(* IEC 61131-3 sources: OpenUnit/plc/projects/GEN/pous/function-blocks, 7 files *)

(* ---- FB_LOOP.st ---- *)
(* PID loop bound to its faceplate tags (<loop>_PV/_SP/_OUT/_MODE/_KP/_TI/_TD/_CSP/_STS).
   Ideal (ISA) PID working in % of span, back-calculation anti-windup, derivative on
   measurement with a 0.1*TD filter, feed-forward and bumpless MAN/AUTO/CAS transfer.
   MODE: 0 MAN, 1 AUTO, 2 CAS.  STS bits: 1 interlock, 2 tracking, 4 high limit, 8 low limit,
   16 cascade setpoint available.  Mirrors Loop + PID in the JavaScript controller runtime. *)
FUNCTION_BLOCK FB_LOOP
  VAR_INPUT
    PV_IN : REAL;              (* process value, engineering units *)
    CSP_IN : REAL;             (* cascade / remote setpoint *)
    CSP_OK : BOOL;             (* remote setpoint supplied and available *)
    FF : REAL;                 (* feed-forward, output engineering units *)
    FORCE_MAN : BOOL;          (* interlock: force manual *)
    TRK : BOOL;                (* track TRK_VAL *)
    TRK_VAL : REAL;
    OUT_HI : REAL := 1.0E30;   (* dynamic output limits, engineering units *)
    OUT_LO : REAL := -1.0E30;
    SP_LO : REAL := -1.0E30;
    SP_HI : REAL := 1.0E30;
    DTS : REAL;                (* simulation time step, s *)
    RESYNC : BOOL;             (* first scan after start-up / initial condition *)
    PV_MIN : REAL := 0.0;      (* configuration from the register map *)
    PV_MAX : REAL := 100.0;
    OUT_MIN : REAL := 0.0;
    OUT_MAX : REAL := 100.0;
    DIRECT : BOOL;             (* direct acting: output rises when PV > SP *)
    SP_TRACK : BOOL := TRUE;   (* setpoint tracks PV in manual *)
    CAS_CFG : BOOL;            (* loop has a cascade input *)
    REF_DT : REAL;             (* > 0: detune when the step exceeds REF_DT (fast time) *)
  END_VAR
  VAR_IN_OUT
    SP : REAL;
    OUT : REAL;
    MODE : DINT;
    KP : REAL;
    TI : REAL;
    TD : REAL;
    PV : REAL;
    CSP : REAL;
    STS : DINT;
  END_VAR
  VAR_OUTPUT
    Q : REAL;                  (* output, engineering units *)
    AUTO : BOOL;               (* not in manual *)
  END_VAR
  VAR
    integ : REAL;
    outPct : REAL;
    prevPv : REAL;
    havePrev : BOOL;
    dState : REAL;
    lastMode : DINT;
    wasTracking : BOOL;
    slow : REAL;
    kpE : REAL;
    tiE : REAL;
    tdE : REAL;
    m : DINT;
    stsW : DINT;
    casOk : BOOL;
    spv : REAL;
    spanO : REAL;
    spanP : REAL;
    ffPct : REAL;
    hiPct : REAL;
    loPct : REAL;
    err : REAL;
    trkPct : REAL;
    p : REAL;
    d : REAL;
    dpv : REAL;
    raw : REAL;
    alpha : REAL;
    hi : REAL;
    lo : REAL;
    unc : REAL;
    doTrack : BOOL;
  END_VAR

  slow := 1.0;
  IF REF_DT > 0.0 AND DTS > REF_DT THEN
    slow := REF_DT / DTS;
  END_IF;
  kpE := MAX(0.0, KP) * slow;
  tiE := MAX(0.0, TI) / slow;
  tdE := MAX(0.0, TD);

  m := MODE;
  IF m > 2 OR m < 0 THEN
    m := 0;
  END_IF;
  stsW := 0;
  IF FORCE_MAN THEN
    m := 0;
    stsW := stsW + 1;
  END_IF;
  casOk := CAS_CFG AND CSP_OK;
  IF casOk THEN
    stsW := stsW + 16;
  END_IF;
  IF m = 2 AND NOT casOk THEN
    m := 1;
  END_IF;
  spv := SP;
  IF m = 2 THEN
    spv := CSP_IN;
  END_IF;
  spv := LIMIT(SP_LO, spv, SP_HI);

  spanO := OUT_MAX - OUT_MIN;
  IF spanO = 0.0 THEN
    spanO := 1.0;
  END_IF;
  spanP := PV_MAX - PV_MIN;
  IF spanP = 0.0 THEN
    spanP := 1.0;
  END_IF;
  ffPct := FF / spanO * 100.0;
  hiPct := 100.0;
  IF OUT_HI < 1.0E29 THEN
    hiPct := (MIN(OUT_HI, OUT_MAX) - OUT_MIN) / spanO * 100.0;
  END_IF;
  loPct := 0.0;
  IF OUT_LO > -1.0E29 THEN
    loPct := (MAX(OUT_LO, OUT_MIN) - OUT_MIN) / spanO * 100.0;
  END_IF;
  err := (spv - PV_IN) / spanP * 100.0;
  IF DIRECT THEN
    err := -err;
  END_IF;

  (* Tracking / manual: force the output and back-calculate the integrator *)
  doTrack := FALSE;
  IF TRK THEN
    trkPct := (TRK_VAL - OUT_MIN) / spanO * 100.0;
    doTrack := TRUE;
    stsW := stsW + 2;
  ELSIF m = 0 THEN
    trkPct := LIMIT(loPct, (OUT - OUT_MIN) / spanO * 100.0, hiPct);
    doTrack := TRUE;
  ELSIF RESYNC OR lastMode = 0 OR wasTracking THEN
    trkPct := (OUT - OUT_MIN) / spanO * 100.0;
    doTrack := TRUE;
  END_IF;
  IF doTrack THEN
    outPct := LIMIT(0.0, trkPct, 100.0);
    integ := outPct - kpE * err - ffPct;
    prevPv := PV_IN;
    havePrev := TRUE;
    dState := 0.0;
  END_IF;

  IF TRK THEN
    IF m = 0 AND SP_TRACK THEN
      spv := PV_IN;
    END_IF;
  ELSIF m = 0 THEN
    IF SP_TRACK THEN
      spv := LIMIT(SP_LO, PV_IN, SP_HI);
    END_IF;
  ELSE
    (* Automatic: PID update *)
    IF DTS > 0.0 THEN
      p := kpE * err;
      IF tiE > 0.0 THEN
        integ := integ + kpE * err * DTS / tiE;
      END_IF;
      d := 0.0;
      IF tdE > 0.0 AND havePrev THEN
        dpv := ((PV_IN - prevPv) / spanP * 100.0) / DTS;
        IF DIRECT THEN
          raw := kpE * tdE * dpv;
        ELSE
          raw := -kpE * tdE * dpv;
        END_IF;
        alpha := DTS / (0.1 * tdE + DTS);
        dState := dState + alpha * (raw - dState);
        d := dState;
      END_IF;
      prevPv := PV_IN;
      havePrev := TRUE;
      hi := MIN(hiPct, 100.0);
      lo := MAX(loPct, 0.0);
      unc := p + integ + d + ffPct;
      outPct := LIMIT(lo, unc, hi);
      IF unc <> outPct THEN
        integ := outPct - p - d - ffPct;
      END_IF;
      IF tiE <= 0.0 THEN
        integ := LIMIT(-1.0E6, integ, 1.0E6);
      END_IF;
    END_IF;
    IF outPct >= hiPct - 0.000001 THEN
      stsW := stsW + 4;
    END_IF;
    IF outPct <= loPct + 0.000001 THEN
      stsW := stsW + 8;
    END_IF;
  END_IF;

  wasTracking := TRK;
  Q := OUT_MIN + outPct / 100.0 * spanO;
  PV := PV_IN;
  SP := spv;
  OUT := Q;
  MODE := m;
  IF CSP_OK THEN
    CSP := CSP_IN;
  ELSE
    CSP := spv;
  END_IF;
  STS := stsW;
  lastMode := m;
  AUTO := m <> 0;
END_FUNCTION_BLOCK

(* ---- FB_MOTOR.st ---- *)
(* Motor / pump / fan device block.  Drives the field command from START/STOP pulses
   (cleared after use), auto start/stop logic and the protective interlock.  A trip of the
   drive is latched (TRIP) until the operator presses STOP, so a standby unit can start on it.
   SYNC (initial condition) aligns the command with the running feedback.  CMD_SET forces the
   command from a sequence, like an operator start without the permissive check. *)
FUNCTION_BLOCK FB_MOTOR
  VAR_INPUT
    RUN_FB : BOOL;             (* field: running *)
    TRIP_FB : BOOL;            (* field: tripped *)
    PERMIT : BOOL := TRUE;     (* start permissive *)
    ILK : BOOL;                (* protective interlock (stops and blocks) *)
    AUTO_START : BOOL;
    AUTO_STOP : BOOL;
    SYNC : BOOL;
    CMD_SET : BOOL;
    CMD_VAL : BOOL;
  END_VAR
  VAR_IN_OUT
    START : BOOL;              (* operator pulse *)
    STOP : BOOL;               (* operator pulse *)
    MODE : DINT;               (* 0 MAN, 1 AUTO / standby *)
    CMD : BOOL;                (* field command *)
    RUN : BOOL;
    TRIP : BOOL;
    PERM : BOOL;
    ILK_T : BOOL;
  END_VAR
  VAR_OUTPUT
    RUNNING : BOOL;
    LATCHED : BOOL;            (* trip latch (cleared by STOP) *)
    TRIPPED : BOOL;            (* field trip or latched trip *)
    IS_AUTO : BOOL;
    REJECTED : BOOL;           (* last start request refused *)
  END_VAR
  VAR
    cmdS : BOOL;
    tripS : BOOL;
  END_VAR

  IF SYNC THEN
    cmdS := RUN_FB;
    tripS := FALSE;
  END_IF;
  IF CMD_SET THEN
    cmdS := CMD_VAL;
    IF CMD_VAL THEN
      tripS := FALSE;
    END_IF;
  END_IF;
  IS_AUTO := MODE = 1;
  IF TRIP_FB THEN
    cmdS := FALSE;
    tripS := TRUE;
  END_IF;
  IF STOP THEN
    cmdS := FALSE;
    tripS := FALSE;
  END_IF;
  IF START THEN
    IF PERMIT AND NOT ILK AND NOT TRIP_FB THEN
      cmdS := TRUE;
      tripS := FALSE;
      REJECTED := FALSE;
    ELSE
      REJECTED := TRUE;
    END_IF;
  END_IF;
  IF IS_AUTO AND AUTO_START AND PERMIT AND NOT ILK AND NOT TRIP_FB AND NOT tripS THEN
    cmdS := TRUE;
  END_IF;
  IF IS_AUTO AND AUTO_STOP THEN
    cmdS := FALSE;
  END_IF;
  IF ILK THEN
    cmdS := FALSE;
  END_IF;
  START := FALSE;
  STOP := FALSE;
  CMD := cmdS;
  RUN := RUN_FB;
  TRIP := tripS;
  PERM := PERMIT;
  ILK_T := ILK;
  RUNNING := RUN_FB;
  LATCHED := tripS;
  TRIPPED := TRIP_FB OR tripS;
END_FUNCTION_BLOCK

(* ---- FB_ONOFF.st ---- *)
(* On/off valve or breaker device block (<dev>_OPEN/_CLOSE pulses, _MODE, _OPENED/_CLOSED,
   _PERM, _ILK).  ILK_OPEN / ILK_CLOSE are protective interlocks; RESET_ON_LOSS drops the
   command when the device leaves the open position by itself (e.g. a breaker trip). *)
FUNCTION_BLOCK FB_ONOFF
  VAR_INPUT
    OPENED_FB : BOOL;          (* field: open / closed position *)
    CLOSED_FB : BOOL;
    HAS_CLOSED : BOOL;         (* a separate closed limit switch exists *)
    PERMIT : BOOL := TRUE;     (* open permissive *)
    CLOSE_PERMIT : BOOL := TRUE;
    ILK_CLOSE : BOOL;
    ILK_OPEN : BOOL;
    AUTO_OPEN : BOOL;
    AUTO_CLOSE : BOOL;
    RESET_ON_LOSS : BOOL;
    SYNC : BOOL;
    CMD_SET : BOOL;
    CMD_VAL : BOOL;
  END_VAR
  VAR_IN_OUT
    OPEN : BOOL;               (* operator pulse *)
    CLOSE : BOOL;              (* operator pulse *)
    MODE : DINT;
    CMD : BOOL;                (* field command *)
    OPENED : BOOL;
    CLOSED : BOOL;
    PERM : BOOL;
    ILK : BOOL;
  END_VAR
  VAR_OUTPUT
    IS_OPEN : BOOL;
    IS_CLOSED : BOOL;
    Q_CMD : BOOL;
    REJECTED : BOOL;
  END_VAR
  VAR
    cmdS : BOOL;
    was : BOOL;
    autoM : BOOL;
  END_VAR

  IF SYNC THEN
    cmdS := OPENED_FB;
    was := OPENED_FB;
  END_IF;
  IF CMD_SET THEN
    cmdS := CMD_VAL;
  END_IF;
  IS_OPEN := OPENED_FB;
  IF HAS_CLOSED THEN
    IS_CLOSED := CLOSED_FB;
  ELSE
    IS_CLOSED := NOT OPENED_FB;
  END_IF;
  autoM := MODE = 1;
  IF RESET_ON_LOSS AND cmdS AND was AND NOT OPENED_FB THEN
    cmdS := FALSE;
  END_IF;
  IF OPEN THEN
    IF PERMIT AND NOT ILK_CLOSE THEN
      cmdS := TRUE;
      REJECTED := FALSE;
    ELSE
      REJECTED := TRUE;
    END_IF;
  END_IF;
  IF CLOSE THEN
    IF CLOSE_PERMIT THEN
      cmdS := FALSE;
      REJECTED := FALSE;
    ELSE
      REJECTED := TRUE;
    END_IF;
  END_IF;
  IF autoM AND AUTO_OPEN AND PERMIT AND NOT ILK_CLOSE THEN
    cmdS := TRUE;
  END_IF;
  IF autoM AND AUTO_CLOSE THEN
    cmdS := FALSE;
  END_IF;
  IF ILK_OPEN THEN
    cmdS := TRUE;
  END_IF;
  IF ILK_CLOSE THEN
    cmdS := FALSE;
  END_IF;
  was := OPENED_FB;
  OPEN := FALSE;
  CLOSE := FALSE;
  CMD := cmdS;
  OPENED := IS_OPEN;
  CLOSED := IS_CLOSED;
  PERM := PERMIT;
  ILK := ILK_CLOSE OR ILK_OPEN;
  Q_CMD := cmdS;
END_FUNCTION_BLOCK

(* ---- FB_PLC_RUNTIME.st ---- *)
(* Controller runtime services, called first in every scan:
   - simulation time step DTS from the plant clock (SIM_TIME_MS), so freeze and fast time
     are honoured by every timer, ramp and PID;
   - initial-condition (IC) commands from the I/O bridge: a new IC_SEQ makes IC_INIT TRUE for
     one scan, the program then resets its internal state; IC_BUILTIN asks for the built-in
     defaults (no snapshot was restored).  The command is acknowledged in IC_ACK;
   - heartbeat, scan counter and a 6 s grace period after start-up / IC load.
   READY stays FALSE until the bridge has initialised the controller once. *)
FUNCTION_BLOCK FB_PLC_RUNTIME
  VAR_INPUT
    SIM_MS : UDINT;            (* plant simulation clock, ms *)
    IC_SEQ : DINT;             (* IC command sequence from the bridge *)
    IC_ID : DINT;              (* IC number *)
    IC_SNAP : BOOL;            (* controller values were restored from a snapshot *)
    CYCLE_MS : REAL := 50.0;   (* task interval, for SCAN_MS *)
  END_VAR
  VAR_IN_OUT
    HEARTBEAT : DINT;
    SCAN_COUNT : UDINT;
    SCAN_MS : REAL;
    SIM_DT : REAL;
    IC_APPLIED : DINT;
    IC_ACK : DINT;
  END_VAR
  VAR_OUTPUT
    DTS : REAL;
    IC_INIT : BOOL;
    IC_BUILTIN : BOOL;
    RESYNC : BOOL;
    GRACE : BOOL;
    READY : BOOL;
  END_VAR
  VAR
    prevMs : UDINT;
    havePrev : BOOL;
    lastSeq : DINT;
    first : BOOL := TRUE;
    graceTmr : TON;
  END_VAR

  (* simulation time step *)
  DTS := 0.0;
  IF havePrev THEN
    DTS := UDINT_TO_REAL(SIM_MS - prevMs) / 1000.0;
    IF DTS < 0.0 OR DTS > 5.0 THEN
      DTS := 0.0;
    END_IF;
  END_IF;
  prevMs := SIM_MS;
  havePrev := TRUE;
  SIM_DT := DTS;

  (* initial condition command *)
  IC_INIT := FALSE;
  IF IC_SEQ <> lastSeq AND IC_SEQ <> 0 THEN
    lastSeq := IC_SEQ;
    IC_INIT := TRUE;
    IC_APPLIED := IC_ID;
    IC_ACK := IC_SEQ;
  END_IF;
  IC_BUILTIN := IC_INIT AND NOT IC_SNAP;
  READY := IC_ACK <> 0;
  RESYNC := IC_INIT OR first;
  first := FALSE;

  graceTmr(IN := NOT IC_INIT, PT := T#6s);
  GRACE := NOT graceTmr.Q;

  HEARTBEAT := HEARTBEAT + 1;
  IF HEARTBEAT > 65535 THEN
    HEARTBEAT := 0;
  END_IF;
  SCAN_COUNT := SCAN_COUNT + 1;
  SCAN_MS := CYCLE_MS;
END_FUNCTION_BLOCK

(* ---- FB_RAMP.st ---- *)
(* Ramp generator: OUT moves towards TARGET at RATE units/s (simulation time).
   INIT loads INIT_VAL (initial condition / bumpless start). *)
FUNCTION_BLOCK FB_RAMP
  VAR_INPUT
    TARGET : REAL;
    RATE : REAL;
    DTS : REAL;
    INIT : BOOL;
    INIT_VAL : REAL;
  END_VAR
  VAR_OUTPUT
    OUT : REAL;
  END_VAR
  VAR
    stepV : REAL;
  END_VAR
  IF INIT THEN
    OUT := INIT_VAL;
  END_IF;
  stepV := RATE * DTS;
  OUT := OUT + LIMIT(-stepV, TARGET - OUT, stepV);
END_FUNCTION_BLOCK

(* ---- FB_STATION.st ---- *)
(* Manual / auto loading station (<station>_OUT/_MODE/_BIAS/_IN/_FB/_STS).
   AUTO: output = auto demand + bias; the bias is computed on the transfer to AUTO so the
   change is bumpless.  STS bits: 1 interlock (forced manual), 2 tracking.
   INIT (initial condition) forgets the previous mode, so a station found in AUTO recomputes
   its bias; with INIT_KEEP (values restored from a snapshot) the bias is kept.  JOIN puts the
   station in AUTO on the master demand with zero bias (auto-started standby unit). *)
FUNCTION_BLOCK FB_STATION
  VAR_INPUT
    AUTO_IN : REAL;            (* auto demand *)
    FB_IN : REAL;              (* position feedback, for display *)
    FORCE_MAN : BOOL;
    TRK : BOOL;
    TRK_VAL : REAL;
    LO : REAL := -1.0E30;      (* output limits; default = station range *)
    HI : REAL := 1.0E30;
    RATE : REAL := 1.0E30;     (* rate limit in AUTO, units/s *)
    DTS : REAL;
    INIT : BOOL;               (* initial condition *)
    INIT_KEEP : BOOL;          (* ... keep the bias (values came from a snapshot) *)
    JOIN : BOOL;               (* go to AUTO with zero bias *)
    OUT_MIN : REAL := 0.0;
    OUT_MAX : REAL := 100.0;
  END_VAR
  VAR_IN_OUT
    OUT : REAL;
    MODE : DINT;
    BIAS : REAL;
    IN_TAG : REAL;
    FB_TAG : REAL;
    STS : DINT;
  END_VAR
  VAR_OUTPUT
    Q : REAL;
    AUTO : BOOL;
  END_VAR
  VAR
    prevMode : DINT;
    m : DINT;
    stsW : DINT;
    cur : REAL;
    o : REAL;
    lo2 : REAL;
    hi2 : REAL;
  END_VAR

  IF INIT THEN
    IF INIT_KEEP AND MODE = 1 THEN
      prevMode := 1;
    ELSE
      prevMode := 0;
    END_IF;
  END_IF;
  IF JOIN THEN
    MODE := 1;
    BIAS := 0.0;
    prevMode := 1;
  END_IF;
  m := 0;
  IF MODE = 1 THEN
    m := 1;
  END_IF;
  stsW := 0;
  IF FORCE_MAN THEN
    m := 0;
    stsW := 1;
  END_IF;
  cur := OUT;
  IF TRK THEN
    o := TRK_VAL;
    stsW := stsW + 2;
  ELSIF m = 1 THEN
    IF prevMode <> 1 THEN
      BIAS := LIMIT(-50.0, cur - AUTO_IN, 50.0);
    END_IF;
    o := AUTO_IN + BIAS;
    IF RATE < 1.0E29 THEN
      o := cur + LIMIT(-RATE * DTS, o - cur, RATE * DTS);
    END_IF;
  ELSE
    o := cur;
  END_IF;
  lo2 := OUT_MIN;
  IF LO > -1.0E29 THEN
    lo2 := LO;
  END_IF;
  hi2 := OUT_MAX;
  IF HI < 1.0E29 THEN
    hi2 := HI;
  END_IF;
  o := LIMIT(lo2, o, hi2);
  prevMode := m;
  OUT := o;
  MODE := m;
  IN_TAG := AUTO_IN;
  FB_TAG := FB_IN;
  STS := stsW;
  Q := o;
  AUTO := m = 1;
END_FUNCTION_BLOCK

(* ---- FB_TONS.st ---- *)
(* On-delay timer running on SIMULATION time (DTS), so it honours freeze and fast time.
   Q goes TRUE once IN has been TRUE for PT seconds.  ET is the elapsed time (s). *)
FUNCTION_BLOCK FB_TONS
  VAR_INPUT
    IN : BOOL;
    PT : REAL;                 (* preset, s *)
    DTS : REAL;
    INIT : BOOL;
  END_VAR
  VAR_OUTPUT
    Q : BOOL;
    ET : REAL;
  END_VAR
  IF INIT THEN
    ET := 0.0;
  END_IF;
  IF IN THEN
    ET := MIN(PT, ET + DTS);
  ELSE
    ET := 0.0;
  END_IF;
  Q := IN AND ET >= PT;
END_FUNCTION_BLOCK
